// Contains tests that verify the XmlControl function block methods
FUNCTION_BLOCK FB_TestXmlControl EXTENDS TcUnit.FB_TestSuite
VAR
    Buffer: ARRAY[0..TcUnit.GVL_Param_TcUnit.xUnitBufferSize - 1] OF BYTE;
END_VAR

Test_NewTag();
Test_NewTagNested();
Test_NewParameter();
Test_NewComment();
Test_CloseOpenTag();
Test_CloseTag();
Test_NewTagData();

METHOD PRIVATE Setup
// Clear buffer
MEMSET(ADR(Buffer), 0, SIZEOF(Buffer));
END_METHOD

METHOD PRIVATE Test_CloseOpenTag
VAR
    XmlControl : FB_XmlControl;
    TagName : STRING := 'MyTag';
    ExpectedBuffer : STRING := '<MyTag/>';
    ActualBuffer : STRING;
    ExpectedResult : STRING;
    ActualResult : STRING;
END_VAR
TEST('Test_CloseOpenTag');

Setup();

XmlControl.SetBuffer(ADR(Buffer), SIZEOF(Buffer));
XmlControl.NewTag(TagName);
XmlControl.CloseTag();
MEMCPY(ADR(ActualBuffer), ADR(Buffer), SIZEOF(ActualBuffer));

AssertEquals_String(Expected := ExpectedBuffer,
                    Actual :=  ActualBuffer,
                    Message := 'Buffer does not contain expected content');

AssertEquals_String(Expected := ExpectedResult,
                    Actual :=  ActualResult,
                    Message := 'CloseTag result does not contain expected content');

TEST_FINISHED();
END_METHOD

METHOD PRIVATE Test_CloseTag
VAR
    XmlControl : FB_XmlControl;
    TagName : STRING := 'MyTag';
    ExpectedBuffer : STRING := '<MyTag>TagData</MyTag>';
    ActualBuffer : STRING;
    ExpectedResult : STRING := '/MyTag';
    ActualResult : STRING;
END_VAR
TEST('Test_CloseTag');

Setup();

XmlControl.SetBuffer(ADR(Buffer), SIZEOF(Buffer));
XmlControl.NewTag(TagName);
XmlControl.NewTagData('TagData');
ActualResult := XmlControl.CloseTag();
MEMCPY(ADR(ActualBuffer), ADR(Buffer), SIZEOF(ActualBuffer));

AssertEquals_String(Expected := ExpectedBuffer,
                    Actual :=  ActualBuffer,
                    Message := 'Buffer does not contain expected content');

AssertEquals_String(Expected := ExpectedResult,
                    Actual :=  ActualResult,
                    Message := 'CloseTag result does not contain expected content');
                   
TEST_FINISHED();
END_METHOD

METHOD PRIVATE Test_NewComment
VAR
    XmlControl : FB_XmlControl;
    Comment : STRING := 'MyComment';
    ExpectedBuffer : STRING := '<!-- MyComment -->';
    ActualBuffer : STRING;
END_VAR
TEST('Test_NewComment');

Setup();

XmlControl.SetBuffer(ADR(Buffer), SIZEOF(Buffer));
XmlControl.NewComment(Comment);
MEMCPY(ADR(ActualBuffer), ADR(Buffer), SIZEOF(ActualBuffer));

AssertEquals_String(Expected := ExpectedBuffer,
                    Actual :=  ActualBuffer,
                    Message := 'Buffer does not contain expected content');

TEST_FINISHED();
END_METHOD

METHOD PRIVATE Test_NewParameter
VAR
    XmlControl : FB_XmlControl;
    XmlEscaped : FB_XmlControl;
    XmlEmpty : FB_XmlControl;
    XmlAdjacent : FB_XmlControl;
    XmlFull : FB_XmlControl;
    XmlLongEscaped : FB_XmlControl;
    ParameterName : STRING := 'ParaName';
    ParameterValue : STRING := 'Value';
    ExpectedBuffer : STRING := ' ParaName="Value"';
    ActualBuffer : STRING;
    LongValue : T_MaxString;
    ValueBytes : POINTER TO BYTE;
    BufferBytes : POINTER TO BYTE;
    Index : INT;
    Length : INT;
END_VAR
VAR CONSTANT
    MAX_SCAN : INT := 1999;
    FULL_VALUE_LENGTH : INT := 255;
    LONG_ESCAPED_COUNT : INT := 60;
    LETTER_A : BYTE := 16#61;
    AMPERSAND : BYTE := 16#26;
    QUOTE_BYTE : BYTE := 16#22;
END_VAR
TEST('Test_NewParameter');

Setup();

XmlControl.SetBuffer(ADR(Buffer), SIZEOF(Buffer));
XmlControl.NewParameter(ParameterName, ParameterValue);
MEMCPY(ADR(ActualBuffer), ADR(Buffer), SIZEOF(ActualBuffer));

AssertEquals_String(Expected := ExpectedBuffer,
                    Actual :=  ActualBuffer,
                    Message := 'Buffer does not contain expected content');

(* Attribute values are escaped (failure messages and TEST_SKIPPED reasons; Codex step-1 re-review R10).
   The cases below are part of this test so the suite keeps its method set; native RED/GREEN is T-6. *)
Setup();
XmlEscaped.SetBuffer(ADR(Buffer), SIZEOF(Buffer));
XmlEscaped.NewParameter('P', 'a"b&c<d>e');
MEMCPY(ADR(ActualBuffer), ADR(Buffer), SIZEOF(ActualBuffer));
AssertEquals_String(Expected := ' P="a&quot;b&amp;c&lt;d&gt;e"', Actual := ActualBuffer,
                    Message := 'Quote, ampersand and angle brackets are not escaped');

Setup();
XmlEmpty.SetBuffer(ADR(Buffer), SIZEOF(Buffer));
XmlEmpty.NewParameter('P', '');
MEMCPY(ADR(ActualBuffer), ADR(Buffer), SIZEOF(ActualBuffer));
AssertEquals_String(Expected := ' P=""', Actual := ActualBuffer, Message := 'Empty value is not an empty attribute');

Setup();
XmlAdjacent.SetBuffer(ADR(Buffer), SIZEOF(Buffer));
XmlAdjacent.NewParameter('P', '&&<<');
MEMCPY(ADR(ActualBuffer), ADR(Buffer), SIZEOF(ActualBuffer));
AssertEquals_String(Expected := ' P="&amp;&amp;&lt;&lt;"', Actual := ActualBuffer, Message := 'Adjacent entities are not escaped');

// A full 255-character value is kept whole: ' P="' + 255 + '"' = 260 bytes.
Setup();
ValueBytes := ADR(LongValue);
FOR Index := 0 TO FULL_VALUE_LENGTH - 1 DO
    ValueBytes[Index] := LETTER_A;
END_FOR
ValueBytes[FULL_VALUE_LENGTH] := 0;
XmlFull.SetBuffer(ADR(Buffer), SIZEOF(Buffer));
XmlFull.NewParameter('P', LongValue);
BufferBytes := ADR(Buffer);
Length := 0;
FOR Index := 0 TO MAX_SCAN DO
    IF BufferBytes[Index] = 0 THEN
        EXIT;
    END_IF
    Length := Length + 1;
END_FOR
AssertEquals_INT(Expected := 4 + FULL_VALUE_LENGTH + 1, Actual := Length, Message := 'A 255-character value is truncated');
AssertEquals_BYTE(Expected := QUOTE_BYTE, Actual := BufferBytes[Length - 1], Message := 'A 255-character value is not closed');

// Escaped output longer than 255 characters: 60 ampersands become 300 bytes of entities.
Setup();
FOR Index := 0 TO LONG_ESCAPED_COUNT - 1 DO
    ValueBytes[Index] := AMPERSAND;
END_FOR
ValueBytes[LONG_ESCAPED_COUNT] := 0;
XmlLongEscaped.SetBuffer(ADR(Buffer), SIZEOF(Buffer));
XmlLongEscaped.NewParameter('P', LongValue);
Length := 0;
FOR Index := 0 TO MAX_SCAN DO
    IF BufferBytes[Index] = 0 THEN
        EXIT;
    END_IF
    Length := Length + 1;
END_FOR
AssertEquals_INT(Expected := 4 + 5 * LONG_ESCAPED_COUNT + 1, Actual := Length, Message := 'Escaped output over 255 characters is truncated');
AssertEquals_BYTE(Expected := QUOTE_BYTE, Actual := BufferBytes[Length - 1], Message := 'Long escaped value is not closed');

TEST_FINISHED();
END_METHOD

METHOD PRIVATE Test_NewTag
VAR
    XmlControl : FB_XmlControl;
    TagName : STRING := 'MyTag';
    ExpectedBuffer : STRING := '<MyTag';
    ActualBuffer : STRING;
END_VAR
TEST('Test_NewTag');

Setup();

XmlControl.SetBuffer(ADR(Buffer), SIZEOF(Buffer));
XmlControl.NewTag(TagName);
MEMCPY(ADR(ActualBuffer), ADR(Buffer), SIZEOF(ActualBuffer));

AssertEquals_String(Expected := ExpectedBuffer,
                    Actual :=  ActualBuffer,
                    Message := 'Buffer does not contain expected content');

TEST_FINISHED();
END_METHOD

METHOD PRIVATE Test_NewTagData
VAR
    XmlControl : FB_XmlControl;
    TagName : STRING := 'MyTag';
    ExpectedBuffer : STRING := '<MyTag>TagData';
    ActualBuffer : STRING;
END_VAR
TEST('Test_NewTagData');

Setup();
XmlControl.SetBuffer(ADR(Buffer), SIZEOF(Buffer));
XmlControl.NewTag(TagName);
XmlControl.NewTagData('TagData');

MEMCPY(ADR(ActualBuffer), ADR(Buffer), SIZEOF(ActualBuffer));

AssertEquals_String(Expected := ExpectedBuffer,
                    Actual :=  ActualBuffer,
                    Message := 'Buffer does not contain expected content');

TEST_FINISHED();
END_METHOD

METHOD PRIVATE Test_NewTagNested
VAR
    XmlControl : FB_XmlControl;
    Tag1Name : STRING := 'MyTag1';
    Tag2Name : STRING := 'MyTag2';
    Tag3Name : STRING := 'MyTag3';
    Tag4Name : STRING := 'MyTag4';
    ExpectedBuffer : STRING := '<MyTag1><MyTag2/><MyTag3/><MyTag4/></MyTag1>';
    ActualBuffer : STRING;
END_VAR
TEST('Test_NewTagNested');

Setup();
XmlControl.SetBuffer(ADR(Buffer), SIZEOF(Buffer));

// <MyTag1><MyTag2/><MyTag3/><MyTag4/></MyTag1>
XmlControl.NewTag(Tag1Name);
XmlControl.NewTag(Tag2Name);
XmlControl.CloseTag();
XmlControl.NewTag(Tag3Name);
XmlControl.CloseTag();
XmlControl.NewTag(Tag4Name);
XmlControl.CloseTag();
XmlControl.CloseTag();

MEMCPY(ADR(ActualBuffer), ADR(Buffer), SIZEOF(ActualBuffer));

AssertEquals_String(Expected := ExpectedBuffer,
                    Actual :=  ActualBuffer,
                    Message := 'Buffer does not contain expected content');

TEST_FINISHED();
END_METHOD

END_FUNCTION_BLOCK

(* stored: Version 1.1.0.1
   POU FB_TestXmlControl: Id {363fde2d-bb7b-452f-a760-baf03449eb88}, SpecialFunc None
   Method Setup: Id {a523e726-082a-4e31-bdb5-31f9c8d19f4c}
   Method Test_CloseOpenTag: Id {7b197c98-60c2-43ce-badc-40234f3381a4}
   Method Test_CloseTag: Id {86a45281-5940-451a-893d-0b71e25ee014}
   Method Test_NewComment: Id {ab168c91-bfbc-487b-89f0-c1ac5f41d253}
   Method Test_NewParameter: Id {284909d6-3d4c-4d69-a860-e3305f25c350}
   Method Test_NewTag: Id {9b9a0770-0e6c-4cd6-899b-75d9d6644278}
   Method Test_NewTagData: Id {3fa16241-ed1c-41c3-a210-bb00b57ea42c}
   Method Test_NewTagNested: Id {127a0665-e103-419e-812d-fe0e6e4c808f} *)
